FUNCTION_BLOCK RETRY_SM
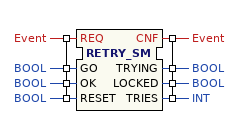
  EVENT_INPUT
    REQ WITH GO, OK, RESET;
  END_EVENT
  EVENT_OUTPUT
    CNF WITH TRYING, LOCKED, TRIES;
  END_EVENT
  VAR_INPUT
    GO : BOOL;
    OK : BOOL;
    RESET : BOOL;
  END_VAR
  VAR_OUTPUT
    TRYING : BOOL;
    LOCKED : BOOL;
    TRIES : INT;
  END_VAR
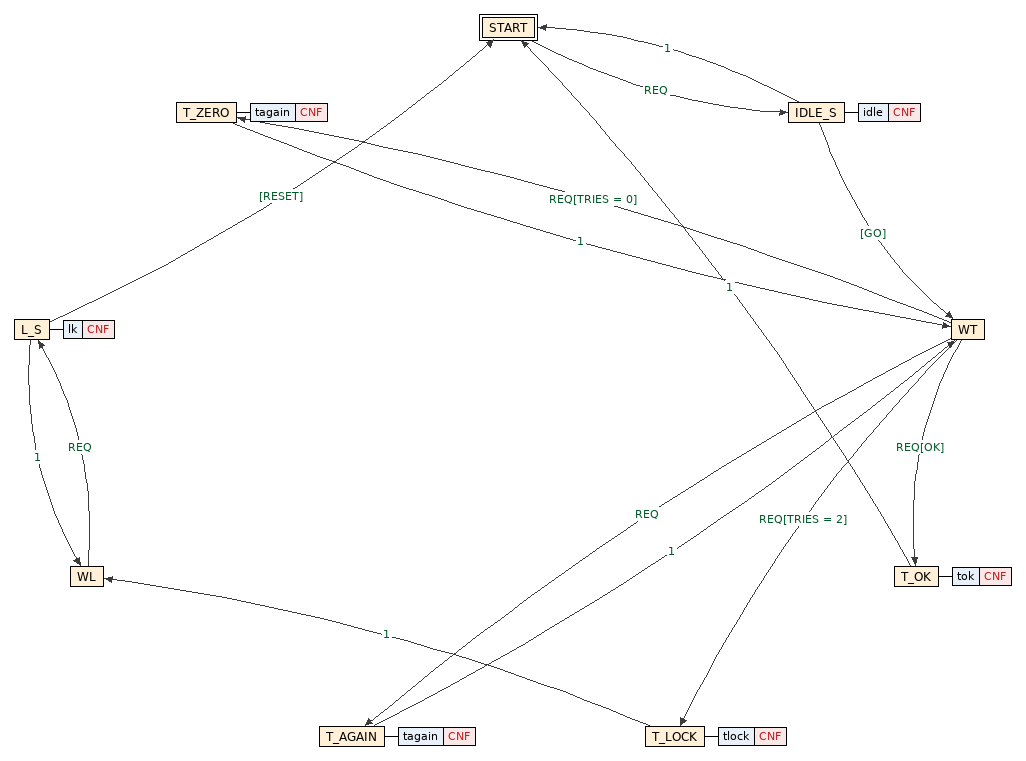
  EC_STATES
    START;
    IDLE_S : idle -> CNF;
    WT;
    T_OK : tok -> CNF;
    T_LOCK : tlock -> CNF;
    T_AGAIN : tagain -> CNF;
    WL;
    L_S : lk -> CNF;
    T_ZERO : tagain -> CNF;
  END_STATES
  EC_TRANSITIONS
    START TO IDLE_S := REQ;
    IDLE_S TO WT := [GO];
    IDLE_S TO START := 1;
    WT TO T_OK := REQ[OK];
    WT TO T_LOCK := REQ[TRIES = 2];
    WT TO T_ZERO := REQ[TRIES = 0];
    WT TO T_AGAIN := REQ;
    T_OK TO START := 1;
    T_LOCK TO WL := 1;
    T_AGAIN TO WT := 1;
    T_ZERO TO WT := 1;
    WL TO L_S := REQ;
    L_S TO START := [RESET];
    L_S TO WL := 1;
  END_TRANSITIONS
  ALGORITHM idle IN ST:
TRYING := FALSE;
TRIES := 0;
  END_ALGORITHM
  ALGORITHM tok IN ST:
TRYING := TRUE;
  END_ALGORITHM
  ALGORITHM tlock IN ST:
TRYING := TRUE;
LOCKED := TRUE;
  END_ALGORITHM
  ALGORITHM tagain IN ST:
TRYING := TRUE;
TRIES := TRIES + 1;
  END_ALGORITHM
  ALGORITHM lk IN ST:
TRYING := FALSE;
IF RESET THEN LOCKED := FALSE; END_IF;
  END_ALGORITHM
END_FUNCTION_BLOCK
